(* IEC 61131-3 sources: BODAS-HelloWorld/st/bodas_rc18_12_40/plc_logic/application/02_easyconfig/dsm_easyconfig/structure (part 3) *)

(* ---- dfc_rbr_ina38scb-DFC_rbr_inA38SCB.st ---- *)
(* --- Interface --- *)
{attribute 'external_name' := 'cmp_rts_DFC_rbr_inA38SCB'}
TYPE DFC_rbr_inA38SCB : STRUCT
		DTC            : UDINT := 16#133100;
		DFCid          : UINT  := 257;
		debounceMethod : USINT := TIME_UP_DOWN;
	END_STRUCT
END_TYPE

(* ---- dfc_rbr_ina38scg-DFC_rbr_inA38SCG.st ---- *)
(* --- Interface --- *)
{attribute 'external_name' := 'cmp_rts_DFC_rbr_inA38SCG'}
TYPE DFC_rbr_inA38SCG : STRUCT
		DTC            : UDINT := 16#133200;
		DFCid          : UINT  := 258;
		debounceMethod : USINT := TIME_UP_DOWN;
	END_STRUCT
END_TYPE

(* ---- dfc_rbr_ina38shuntscb-DFC_rbr_inA38ShuntSCB.st ---- *)
(* --- Interface --- *)
{attribute 'external_name' := 'cmp_rts_DFC_rbr_inA38ShuntSCB'}
TYPE DFC_rbr_inA38ShuntSCB : STRUCT
		DTC            : UDINT := 16#133300;
		DFCid          : UINT  := 259;
		debounceMethod : USINT := TIME_UP_DOWN;
	END_STRUCT
END_TYPE

(* ---- dfc_rbr_ina39aicscb-DFC_rbr_inA39AicSCB.st ---- *)
(* --- Interface --- *)
{attribute 'external_name' := 'cmp_rts_DFC_rbr_inA39AicSCB'}
TYPE DFC_rbr_inA39AicSCB : STRUCT
		DTC            : UDINT := 16#133400;
		DFCid          : UINT  := 260;
		debounceMethod : USINT := TIME_UP_DOWN;
	END_STRUCT
END_TYPE

(* ---- dfc_rbr_ina39aicscg-DFC_rbr_inA39AicSCG.st ---- *)
(* --- Interface --- *)
{attribute 'external_name' := 'cmp_rts_DFC_rbr_inA39AicSCG'}
TYPE DFC_rbr_inA39AicSCG : STRUCT
		DTC            : UDINT := 16#133500;
		DFCid          : UINT  := 261;
		debounceMethod : USINT := TIME_UP_DOWN;
	END_STRUCT
END_TYPE

(* ---- dfc_rbr_ina39or-DFC_rbr_inA39OR.st ---- *)
(* --- Interface --- *)
{attribute 'external_name' := 'cmp_rts_DFC_rbr_inA39OR'}
TYPE DFC_rbr_inA39OR : STRUCT
		DTC            : UDINT := 16#133600;
		DFCid          : UINT  := 262;
		debounceMethod : USINT := TIME_UP_DOWN;
	END_STRUCT
END_TYPE

(* ---- dfc_rbr_ina39scb-DFC_rbr_inA39SCB.st ---- *)
(* --- Interface --- *)
{attribute 'external_name' := 'cmp_rts_DFC_rbr_inA39SCB'}
TYPE DFC_rbr_inA39SCB : STRUCT
		DTC            : UDINT := 16#133700;
		DFCid          : UINT  := 263;
		debounceMethod : USINT := TIME_UP_DOWN;
	END_STRUCT
END_TYPE

(* ---- dfc_rbr_ina39scg-DFC_rbr_inA39SCG.st ---- *)
(* --- Interface --- *)
{attribute 'external_name' := 'cmp_rts_DFC_rbr_inA39SCG'}
TYPE DFC_rbr_inA39SCG : STRUCT
		DTC            : UDINT := 16#133800;
		DFCid          : UINT  := 264;
		debounceMethod : USINT := TIME_UP_DOWN;
	END_STRUCT
END_TYPE

(* ---- dfc_rbr_ina39shuntscb-DFC_rbr_inA39ShuntSCB.st ---- *)
(* --- Interface --- *)
{attribute 'external_name' := 'cmp_rts_DFC_rbr_inA39ShuntSCB'}
TYPE DFC_rbr_inA39ShuntSCB : STRUCT
		DTC            : UDINT := 16#133900;
		DFCid          : UINT  := 265;
		debounceMethod : USINT := TIME_UP_DOWN;
	END_STRUCT
END_TYPE

(* ---- dfc_rbr_ina40or-DFC_rbr_inA40OR.st ---- *)
(* --- Interface --- *)
{attribute 'external_name' := 'cmp_rts_DFC_rbr_inA40OR'}
TYPE DFC_rbr_inA40OR : STRUCT
		DTC            : UDINT := 16#133A00;
		DFCid          : UINT  := 266;
		debounceMethod : USINT := TIME_UP_DOWN;
	END_STRUCT
END_TYPE

(* ---- dfc_rbr_ina40scb-DFC_rbr_inA40SCB.st ---- *)
(* --- Interface --- *)
{attribute 'external_name' := 'cmp_rts_DFC_rbr_inA40SCB'}
TYPE DFC_rbr_inA40SCB : STRUCT
		DTC            : UDINT := 16#133B00;
		DFCid          : UINT  := 267;
		debounceMethod : USINT := TIME_UP_DOWN;
	END_STRUCT
END_TYPE

(* ---- dfc_rbr_ina40scg-DFC_rbr_inA40SCG.st ---- *)
(* --- Interface --- *)
{attribute 'external_name' := 'cmp_rts_DFC_rbr_inA40SCG'}
TYPE DFC_rbr_inA40SCG : STRUCT
		DTC            : UDINT := 16#133C00;
		DFCid          : UINT  := 268;
		debounceMethod : USINT := TIME_UP_DOWN;
	END_STRUCT
END_TYPE

(* ---- dfc_rbr_ina41or-DFC_rbr_inA41OR.st ---- *)
(* --- Interface --- *)
{attribute 'external_name' := 'cmp_rts_DFC_rbr_inA41OR'}
TYPE DFC_rbr_inA41OR : STRUCT
		DTC            : UDINT := 16#133D00;
		DFCid          : UINT  := 269;
		debounceMethod : USINT := TIME_UP_DOWN;
	END_STRUCT
END_TYPE

(* ---- dfc_rbr_ina41scb-DFC_rbr_inA41SCB.st ---- *)
(* --- Interface --- *)
{attribute 'external_name' := 'cmp_rts_DFC_rbr_inA41SCB'}
TYPE DFC_rbr_inA41SCB : STRUCT
		DTC            : UDINT := 16#133E00;
		DFCid          : UINT  := 270;
		debounceMethod : USINT := TIME_UP_DOWN;
	END_STRUCT
END_TYPE

(* ---- dfc_rbr_ina41scg-DFC_rbr_inA41SCG.st ---- *)
(* --- Interface --- *)
{attribute 'external_name' := 'cmp_rts_DFC_rbr_inA41SCG'}
TYPE DFC_rbr_inA41SCG : STRUCT
		DTC            : UDINT := 16#133F00;
		DFCid          : UINT  := 271;
		debounceMethod : USINT := TIME_UP_DOWN;
	END_STRUCT
END_TYPE

(* ---- dfc_rbr_ina42or-DFC_rbr_inA42OR.st ---- *)
(* --- Interface --- *)
{attribute 'external_name' := 'cmp_rts_DFC_rbr_inA42OR'}
TYPE DFC_rbr_inA42OR : STRUCT
		DTC            : UDINT := 16#134000;
		DFCid          : UINT  := 272;
		debounceMethod : USINT := TIME_UP_DOWN;
	END_STRUCT
END_TYPE

(* ---- dfc_rbr_ina42scb-DFC_rbr_inA42SCB.st ---- *)
(* --- Interface --- *)
{attribute 'external_name' := 'cmp_rts_DFC_rbr_inA42SCB'}
TYPE DFC_rbr_inA42SCB : STRUCT
		DTC            : UDINT := 16#134100;
		DFCid          : UINT  := 273;
		debounceMethod : USINT := TIME_UP_DOWN;
	END_STRUCT
END_TYPE

(* ---- dfc_rbr_ina42scg-DFC_rbr_inA42SCG.st ---- *)
(* --- Interface --- *)
{attribute 'external_name' := 'cmp_rts_DFC_rbr_inA42SCG'}
TYPE DFC_rbr_inA42SCG : STRUCT
		DTC            : UDINT := 16#134200;
		DFCid          : UINT  := 274;
		debounceMethod : USINT := TIME_UP_DOWN;
	END_STRUCT
END_TYPE

(* ---- dfc_rbr_ina43aicscb-DFC_rbr_inA43AicSCB.st ---- *)
(* --- Interface --- *)
{attribute 'external_name' := 'cmp_rts_DFC_rbr_inA43AicSCB'}
TYPE DFC_rbr_inA43AicSCB : STRUCT
		DTC            : UDINT := 16#134300;
		DFCid          : UINT  := 275;
		debounceMethod : USINT := TIME_UP_DOWN;
	END_STRUCT
END_TYPE

(* ---- dfc_rbr_ina43aicscg-DFC_rbr_inA43AicSCG.st ---- *)
(* --- Interface --- *)
{attribute 'external_name' := 'cmp_rts_DFC_rbr_inA43AicSCG'}
TYPE DFC_rbr_inA43AicSCG : STRUCT
		DTC            : UDINT := 16#134400;
		DFCid          : UINT  := 276;
		debounceMethod : USINT := TIME_UP_DOWN;
	END_STRUCT
END_TYPE

(* ---- dfc_rbr_ina43or-DFC_rbr_inA43OR.st ---- *)
(* --- Interface --- *)
{attribute 'external_name' := 'cmp_rts_DFC_rbr_inA43OR'}
TYPE DFC_rbr_inA43OR : STRUCT
		DTC            : UDINT := 16#134500;
		DFCid          : UINT  := 277;
		debounceMethod : USINT := TIME_UP_DOWN;
	END_STRUCT
END_TYPE

(* ---- dfc_rbr_ina43scb-DFC_rbr_inA43SCB.st ---- *)
(* --- Interface --- *)
{attribute 'external_name' := 'cmp_rts_DFC_rbr_inA43SCB'}
TYPE DFC_rbr_inA43SCB : STRUCT
		DTC            : UDINT := 16#134600;
		DFCid          : UINT  := 278;
		debounceMethod : USINT := TIME_UP_DOWN;
	END_STRUCT
END_TYPE

(* ---- dfc_rbr_ina43scg-DFC_rbr_inA43SCG.st ---- *)
(* --- Interface --- *)
{attribute 'external_name' := 'cmp_rts_DFC_rbr_inA43SCG'}
TYPE DFC_rbr_inA43SCG : STRUCT
		DTC            : UDINT := 16#134700;
		DFCid          : UINT  := 279;
		debounceMethod : USINT := TIME_UP_DOWN;
	END_STRUCT
END_TYPE

(* ---- dfc_rbr_ina43shuntscb-DFC_rbr_inA43ShuntSCB.st ---- *)
(* --- Interface --- *)
{attribute 'external_name' := 'cmp_rts_DFC_rbr_inA43ShuntSCB'}
TYPE DFC_rbr_inA43ShuntSCB : STRUCT
		DTC            : UDINT := 16#134800;
		DFCid          : UINT  := 280;
		debounceMethod : USINT := TIME_UP_DOWN;
	END_STRUCT
END_TYPE

(* ---- dfc_rbr_ina44ol-DFC_rbr_inA44OL.st ---- *)
(* --- Interface --- *)
{attribute 'external_name' := 'cmp_rts_DFC_rbr_inA44OL'}
TYPE DFC_rbr_inA44OL : STRUCT
		DTC            : UDINT := 16#134900;
		DFCid          : UINT  := 281;
		debounceMethod : USINT := TIME_UP_DOWN;
	END_STRUCT
END_TYPE

(* ---- dfc_rbr_ina44scb-DFC_rbr_inA44SCB.st ---- *)
(* --- Interface --- *)
{attribute 'external_name' := 'cmp_rts_DFC_rbr_inA44SCB'}
TYPE DFC_rbr_inA44SCB : STRUCT
		DTC            : UDINT := 16#134A00;
		DFCid          : UINT  := 282;
		debounceMethod : USINT := TIME_UP_DOWN;
	END_STRUCT
END_TYPE

(* ---- dfc_rbr_ina44scg-DFC_rbr_inA44SCG.st ---- *)
(* --- Interface --- *)
{attribute 'external_name' := 'cmp_rts_DFC_rbr_inA44SCG'}
TYPE DFC_rbr_inA44SCG : STRUCT
		DTC            : UDINT := 16#134B00;
		DFCid          : UINT  := 283;
		debounceMethod : USINT := TIME_UP_DOWN;
	END_STRUCT
END_TYPE

(* ---- dfc_rbr_ina57or-DFC_rbr_inA57OR.st ---- *)
(* --- Interface --- *)
{attribute 'external_name' := 'cmp_rts_DFC_rbr_inA57OR'}
TYPE DFC_rbr_inA57OR : STRUCT
		DTC            : UDINT := 16#134C00;
		DFCid          : UINT  := 284;
		debounceMethod : USINT := TIME_UP_DOWN;
	END_STRUCT
END_TYPE

(* ---- dfc_rbr_ina57scb-DFC_rbr_inA57SCB.st ---- *)
(* --- Interface --- *)
{attribute 'external_name' := 'cmp_rts_DFC_rbr_inA57SCB'}
TYPE DFC_rbr_inA57SCB : STRUCT
		DTC            : UDINT := 16#134D00;
		DFCid          : UINT  := 285;
		debounceMethod : USINT := TIME_UP_DOWN;
	END_STRUCT
END_TYPE

(* ---- dfc_rbr_ina57scg-DFC_rbr_inA57SCG.st ---- *)
(* --- Interface --- *)
{attribute 'external_name' := 'cmp_rts_DFC_rbr_inA57SCG'}
TYPE DFC_rbr_inA57SCG : STRUCT
		DTC            : UDINT := 16#134E00;
		DFCid          : UINT  := 286;
		debounceMethod : USINT := TIME_UP_DOWN;
	END_STRUCT
END_TYPE

(* ---- dfc_rbr_ina59ol-DFC_rbr_inA59OL.st ---- *)
(* --- Interface --- *)
{attribute 'external_name' := 'cmp_rts_DFC_rbr_inA59OL'}
TYPE DFC_rbr_inA59OL : STRUCT
		DTC            : UDINT := 16#134F00;
		DFCid          : UINT  := 287;
		debounceMethod : USINT := TIME_UP_DOWN;
	END_STRUCT
END_TYPE

(* ---- dfc_rbr_ina59scb-DFC_rbr_inA59SCB.st ---- *)
(* --- Interface --- *)
{attribute 'external_name' := 'cmp_rts_DFC_rbr_inA59SCB'}
TYPE DFC_rbr_inA59SCB : STRUCT
		DTC            : UDINT := 16#135000;
		DFCid          : UINT  := 288;
		debounceMethod : USINT := TIME_UP_DOWN;
	END_STRUCT
END_TYPE

(* ---- dfc_rbr_ina59scg-DFC_rbr_inA59SCG.st ---- *)
(* --- Interface --- *)
{attribute 'external_name' := 'cmp_rts_DFC_rbr_inA59SCG'}
TYPE DFC_rbr_inA59SCG : STRUCT
		DTC            : UDINT := 16#135100;
		DFCid          : UINT  := 289;
		debounceMethod : USINT := TIME_UP_DOWN;
	END_STRUCT
END_TYPE

(* ---- dfc_rbr_inai-DFC_rbr_inAi.st ---- *)
(* --- Interface --- *)
{attribute 'external_name' := 'cmp_rts_DFC_rbr_inAi'}
TYPE DFC_rbr_inAi : STRUCT
		DTC            : UDINT := 16#038000;
		DFCid          : UINT  := 882;
		debounceMethod : USINT := NO_DEBOUNCE;
	END_STRUCT
END_TYPE

(* ---- dfc_rbr_inaic-DFC_rbr_inAic.st ---- *)
(* --- Interface --- *)
{attribute 'external_name' := 'cmp_rts_DFC_rbr_inAic'}
TYPE DFC_rbr_inAic : STRUCT
		DTC            : UDINT := 16#038100;
		DFCid          : UINT  := 883;
		debounceMethod : USINT := NO_DEBOUNCE;
	END_STRUCT
END_TYPE

(* ---- dfc_rbr_inaiccfg-DFC_rbr_inAicCfg.st ---- *)
(* --- Interface --- *)
{attribute 'external_name' := 'cmp_rts_DFC_rbr_inAicCfg'}
TYPE DFC_rbr_inAicCfg : STRUCT
		DTC            : UDINT := 16#038200;
		DFCid          : UINT  := 884;
		debounceMethod : USINT := NO_DEBOUNCE;
	END_STRUCT
END_TYPE

(* ---- dfc_rbr_inaicgetstatus-DFC_rbr_inAicGetStatus.st ---- *)
(* --- Interface --- *)
{attribute 'external_name' := 'cmp_rts_DFC_rbr_inAicGetStatus'}
TYPE DFC_rbr_inAicGetStatus : STRUCT
		DTC            : UDINT := 16#038D00;
		DFCid          : UINT  := 885;
		debounceMethod : USINT := NO_DEBOUNCE;
	END_STRUCT
END_TYPE

(* ---- dfc_rbr_inaid-DFC_rbr_inAid.st ---- *)
(* --- Interface --- *)
{attribute 'external_name' := 'cmp_rts_DFC_rbr_inAid'}
TYPE DFC_rbr_inAid : STRUCT
		DTC            : UDINT := 16#038300;
		DFCid          : UINT  := 886;
		debounceMethod : USINT := NO_DEBOUNCE;
	END_STRUCT
END_TYPE

(* ---- dfc_rbr_inaidcfg-DFC_rbr_inAidCfg.st ---- *)
(* --- Interface --- *)
{attribute 'external_name' := 'cmp_rts_DFC_rbr_inAidCfg'}
TYPE DFC_rbr_inAidCfg : STRUCT
		DTC            : UDINT := 16#038400;
		DFCid          : UINT  := 887;
		debounceMethod : USINT := NO_DEBOUNCE;
	END_STRUCT
END_TYPE

(* ---- dfc_rbr_inaiv-DFC_rbr_inAiv.st ---- *)
(* --- Interface --- *)
{attribute 'external_name' := 'cmp_rts_DFC_rbr_inAiv'}
TYPE DFC_rbr_inAiv : STRUCT
		DTC            : UDINT := 16#038500;
		DFCid          : UINT  := 888;
		debounceMethod : USINT := NO_DEBOUNCE;
	END_STRUCT
END_TYPE

(* ---- dfc_rbr_inaivcfg-DFC_rbr_inAivCfg.st ---- *)
(* --- Interface --- *)
{attribute 'external_name' := 'cmp_rts_DFC_rbr_inAivCfg'}
TYPE DFC_rbr_inAivCfg : STRUCT
		DTC            : UDINT := 16#038600;
		DFCid          : UINT  := 889;
		debounceMethod : USINT := NO_DEBOUNCE;
	END_STRUCT
END_TYPE

(* ---- dfc_rbr_inaivgetstatus-DFC_rbr_inAivGetStatus.st ---- *)
(* --- Interface --- *)
{attribute 'external_name' := 'cmp_rts_DFC_rbr_inAivGetStatus'}
TYPE DFC_rbr_inAivGetStatus : STRUCT
		DTC            : UDINT := 16#038C00;
		DFCid          : UINT  := 890;
		debounceMethod : USINT := NO_DEBOUNCE;
	END_STRUCT
END_TYPE

(* ---- dfc_rbr_indi-DFC_rbr_inDi.st ---- *)
(* --- Interface --- *)
{attribute 'external_name' := 'cmp_rts_DFC_rbr_inDi'}
TYPE DFC_rbr_inDi : STRUCT
		DTC            : UDINT := 16#038700;
		DFCid          : UINT  := 891;
		debounceMethod : USINT := NO_DEBOUNCE;
	END_STRUCT
END_TYPE

(* ---- dfc_rbr_infi-DFC_rbr_inFi.st ---- *)
(* --- Interface --- *)
{attribute 'external_name' := 'cmp_rts_DFC_rbr_inFi'}
TYPE DFC_rbr_inFi : STRUCT
		DTC            : UDINT := 16#038800;
		DFCid          : UINT  := 892;
		debounceMethod : USINT := NO_DEBOUNCE;
	END_STRUCT
END_TYPE

(* ---- dfc_rbr_infi_buffered-DFC_rbr_inFi_Buffered.st ---- *)
(* --- Interface --- *)
{attribute 'external_name' := 'cmp_rts_DFC_rbr_inFi_Buffered'}
TYPE DFC_rbr_inFi_Buffered : STRUCT
		DTC            : UDINT := 16#135200;
		DFCid          : UINT  := 895;
		debounceMethod : USINT := NO_DEBOUNCE;
	END_STRUCT
END_TYPE

(* ---- dfc_rbr_inficfg-DFC_rbr_inFiCfg.st ---- *)
(* --- Interface --- *)
{attribute 'external_name' := 'cmp_rts_DFC_rbr_inFiCfg'}
TYPE DFC_rbr_inFiCfg : STRUCT
		DTC            : UDINT := 16#038900;
		DFCid          : UINT  := 893;
		debounceMethod : USINT := NO_DEBOUNCE;
	END_STRUCT
END_TYPE

(* ---- dfc_rbr_infigetstatus-DFC_rbr_inFiGetStatus.st ---- *)
(* --- Interface --- *)
{attribute 'external_name' := 'cmp_rts_DFC_rbr_inFiGetStatus'}
TYPE DFC_rbr_inFiGetStatus : STRUCT
		DTC            : UDINT := 16#038F00;
		DFCid          : UINT  := 894;
		debounceMethod : USINT := NO_DEBOUNCE;
	END_STRUCT
END_TYPE

(* ---- dfc_rbr_ink10or-DFC_rbr_inK10OR.st ---- *)
(* --- Interface --- *)
{attribute 'external_name' := 'cmp_rts_DFC_rbr_inK10OR'}
TYPE DFC_rbr_inK10OR : STRUCT
		DTC            : UDINT := 16#030100;
		DFCid          : UINT  := 290;
		debounceMethod : USINT := TIME_UP_DOWN;
	END_STRUCT
END_TYPE

(* ---- dfc_rbr_ink10scb-DFC_rbr_inK10SCB.st ---- *)
(* --- Interface --- *)
{attribute 'external_name' := 'cmp_rts_DFC_rbr_inK10SCB'}
TYPE DFC_rbr_inK10SCB : STRUCT
		DTC            : UDINT := 16#030200;
		DFCid          : UINT  := 291;
		debounceMethod : USINT := TIME_UP_DOWN;
	END_STRUCT
END_TYPE

(* ---- dfc_rbr_ink10scg-DFC_rbr_inK10SCG.st ---- *)
(* --- Interface --- *)
{attribute 'external_name' := 'cmp_rts_DFC_rbr_inK10SCG'}
TYPE DFC_rbr_inK10SCG : STRUCT
		DTC            : UDINT := 16#030300;
		DFCid          : UINT  := 292;
		debounceMethod : USINT := TIME_UP_DOWN;
	END_STRUCT
END_TYPE

(* ---- dfc_rbr_ink11or-DFC_rbr_inK11OR.st ---- *)
(* --- Interface --- *)
{attribute 'external_name' := 'cmp_rts_DFC_rbr_inK11OR'}
TYPE DFC_rbr_inK11OR : STRUCT
		DTC            : UDINT := 16#03A200;
		DFCid          : UINT  := 293;
		debounceMethod : USINT := TIME_UP_DOWN;
	END_STRUCT
END_TYPE

(* ---- dfc_rbr_ink11scb-DFC_rbr_inK11SCB.st ---- *)
(* --- Interface --- *)
{attribute 'external_name' := 'cmp_rts_DFC_rbr_inK11SCB'}
TYPE DFC_rbr_inK11SCB : STRUCT
		DTC            : UDINT := 16#03A300;
		DFCid          : UINT  := 294;
		debounceMethod : USINT := TIME_UP_DOWN;
	END_STRUCT
END_TYPE

(* ---- dfc_rbr_ink11scg-DFC_rbr_inK11SCG.st ---- *)
(* --- Interface --- *)
{attribute 'external_name' := 'cmp_rts_DFC_rbr_inK11SCG'}
TYPE DFC_rbr_inK11SCG : STRUCT
		DTC            : UDINT := 16#03A400;
		DFCid          : UINT  := 295;
		debounceMethod : USINT := TIME_UP_DOWN;
	END_STRUCT
END_TYPE

(* ---- dfc_rbr_ink30aicscb-DFC_rbr_inK30AicSCB.st ---- *)
(* --- Interface --- *)
{attribute 'external_name' := 'cmp_rts_DFC_rbr_inK30AicSCB'}
TYPE DFC_rbr_inK30AicSCB : STRUCT
		DTC            : UDINT := 16#03A500;
		DFCid          : UINT  := 296;
		debounceMethod : USINT := TIME_UP_DOWN;
	END_STRUCT
END_TYPE

(* ---- dfc_rbr_ink30aicscg-DFC_rbr_inK30AicSCG.st ---- *)
(* --- Interface --- *)
{attribute 'external_name' := 'cmp_rts_DFC_rbr_inK30AicSCG'}
TYPE DFC_rbr_inK30AicSCG : STRUCT
		DTC            : UDINT := 16#03A600;
		DFCid          : UINT  := 297;
		debounceMethod : USINT := TIME_UP_DOWN;
	END_STRUCT
END_TYPE

(* ---- dfc_rbr_ink30or-DFC_rbr_inK30OR.st ---- *)
(* --- Interface --- *)
{attribute 'external_name' := 'cmp_rts_DFC_rbr_inK30OR'}
TYPE DFC_rbr_inK30OR : STRUCT
		DTC            : UDINT := 16#03A700;
		DFCid          : UINT  := 298;
		debounceMethod : USINT := TIME_UP_DOWN;
	END_STRUCT
END_TYPE

(* ---- dfc_rbr_ink30scb-DFC_rbr_inK30SCB.st ---- *)
(* --- Interface --- *)
{attribute 'external_name' := 'cmp_rts_DFC_rbr_inK30SCB'}
TYPE DFC_rbr_inK30SCB : STRUCT
		DTC            : UDINT := 16#03A800;
		DFCid          : UINT  := 299;
		debounceMethod : USINT := TIME_UP_DOWN;
	END_STRUCT
END_TYPE

(* ---- dfc_rbr_ink30scg-DFC_rbr_inK30SCG.st ---- *)
(* --- Interface --- *)
{attribute 'external_name' := 'cmp_rts_DFC_rbr_inK30SCG'}
TYPE DFC_rbr_inK30SCG : STRUCT
		DTC            : UDINT := 16#03A900;
		DFCid          : UINT  := 300;
		debounceMethod : USINT := TIME_UP_DOWN;
	END_STRUCT
END_TYPE

(* ---- dfc_rbr_ink30shuntscb-DFC_rbr_inK30ShuntSCB.st ---- *)
(* --- Interface --- *)
{attribute 'external_name' := 'cmp_rts_DFC_rbr_inK30ShuntSCB'}
TYPE DFC_rbr_inK30ShuntSCB : STRUCT
		DTC            : UDINT := 16#03AA00;
		DFCid          : UINT  := 301;
		debounceMethod : USINT := TIME_UP_DOWN;
	END_STRUCT
END_TYPE

(* ---- dfc_rbr_ink31or-DFC_rbr_inK31OR.st ---- *)
(* --- Interface --- *)
{attribute 'external_name' := 'cmp_rts_DFC_rbr_inK31OR'}
TYPE DFC_rbr_inK31OR : STRUCT
		DTC            : UDINT := 16#03AB00;
		DFCid          : UINT  := 302;
		debounceMethod : USINT := TIME_UP_DOWN;
	END_STRUCT
END_TYPE

(* ---- dfc_rbr_ink31scb-DFC_rbr_inK31SCB.st ---- *)
(* --- Interface --- *)
{attribute 'external_name' := 'cmp_rts_DFC_rbr_inK31SCB'}
TYPE DFC_rbr_inK31SCB : STRUCT
		DTC            : UDINT := 16#03AC00;
		DFCid          : UINT  := 303;
		debounceMethod : USINT := TIME_UP_DOWN;
	END_STRUCT
END_TYPE

(* ---- dfc_rbr_ink31scg-DFC_rbr_inK31SCG.st ---- *)
(* --- Interface --- *)
{attribute 'external_name' := 'cmp_rts_DFC_rbr_inK31SCG'}
TYPE DFC_rbr_inK31SCG : STRUCT
		DTC            : UDINT := 16#03AD00;
		DFCid          : UINT  := 304;
		debounceMethod : USINT := TIME_UP_DOWN;
	END_STRUCT
END_TYPE

(* ---- dfc_rbr_ink32or-DFC_rbr_inK32OR.st ---- *)
(* --- Interface --- *)
{attribute 'external_name' := 'cmp_rts_DFC_rbr_inK32OR'}
TYPE DFC_rbr_inK32OR : STRUCT
		DTC            : UDINT := 16#03AE00;
		DFCid          : UINT  := 305;
		debounceMethod : USINT := TIME_UP_DOWN;
	END_STRUCT
END_TYPE

(* ---- dfc_rbr_ink32scb-DFC_rbr_inK32SCB.st ---- *)
(* --- Interface --- *)
{attribute 'external_name' := 'cmp_rts_DFC_rbr_inK32SCB'}
TYPE DFC_rbr_inK32SCB : STRUCT
		DTC            : UDINT := 16#03AF00;
		DFCid          : UINT  := 306;
		debounceMethod : USINT := TIME_UP_DOWN;
	END_STRUCT
END_TYPE

(* ---- dfc_rbr_ink32scg-DFC_rbr_inK32SCG.st ---- *)
(* --- Interface --- *)
{attribute 'external_name' := 'cmp_rts_DFC_rbr_inK32SCG'}
TYPE DFC_rbr_inK32SCG : STRUCT
		DTC            : UDINT := 16#03B000;
		DFCid          : UINT  := 307;
		debounceMethod : USINT := TIME_UP_DOWN;
	END_STRUCT
END_TYPE

(* ---- dfc_rbr_ink33or-DFC_rbr_inK33OR.st ---- *)
(* --- Interface --- *)
{attribute 'external_name' := 'cmp_rts_DFC_rbr_inK33OR'}
TYPE DFC_rbr_inK33OR : STRUCT
		DTC            : UDINT := 16#03B100;
		DFCid          : UINT  := 308;
		debounceMethod : USINT := TIME_UP_DOWN;
	END_STRUCT
END_TYPE

(* ---- dfc_rbr_ink33scb-DFC_rbr_inK33SCB.st ---- *)
(* --- Interface --- *)
{attribute 'external_name' := 'cmp_rts_DFC_rbr_inK33SCB'}
TYPE DFC_rbr_inK33SCB : STRUCT
		DTC            : UDINT := 16#03B200;
		DFCid          : UINT  := 309;
		debounceMethod : USINT := TIME_UP_DOWN;
	END_STRUCT
END_TYPE

(* ---- dfc_rbr_ink33scg-DFC_rbr_inK33SCG.st ---- *)
(* --- Interface --- *)
{attribute 'external_name' := 'cmp_rts_DFC_rbr_inK33SCG'}
TYPE DFC_rbr_inK33SCG : STRUCT
		DTC            : UDINT := 16#03B300;
		DFCid          : UINT  := 310;
		debounceMethod : USINT := TIME_UP_DOWN;
	END_STRUCT
END_TYPE

(* ---- dfc_rbr_ink34or-DFC_rbr_inK34OR.st ---- *)
(* --- Interface --- *)
{attribute 'external_name' := 'cmp_rts_DFC_rbr_inK34OR'}
TYPE DFC_rbr_inK34OR : STRUCT
		DTC            : UDINT := 16#03B400;
		DFCid          : UINT  := 311;
		debounceMethod : USINT := TIME_UP_DOWN;
	END_STRUCT
END_TYPE

(* ---- dfc_rbr_ink34scb-DFC_rbr_inK34SCB.st ---- *)
(* --- Interface --- *)
{attribute 'external_name' := 'cmp_rts_DFC_rbr_inK34SCB'}
TYPE DFC_rbr_inK34SCB : STRUCT
		DTC            : UDINT := 16#03B500;
		DFCid          : UINT  := 312;
		debounceMethod : USINT := TIME_UP_DOWN;
	END_STRUCT
END_TYPE

(* ---- dfc_rbr_ink34scg-DFC_rbr_inK34SCG.st ---- *)
(* --- Interface --- *)
{attribute 'external_name' := 'cmp_rts_DFC_rbr_inK34SCG'}
TYPE DFC_rbr_inK34SCG : STRUCT
		DTC            : UDINT := 16#03B600;
		DFCid          : UINT  := 313;
		debounceMethod : USINT := TIME_UP_DOWN;
	END_STRUCT
END_TYPE

(* ---- dfc_rbr_ink35or-DFC_rbr_inK35OR.st ---- *)
(* --- Interface --- *)
{attribute 'external_name' := 'cmp_rts_DFC_rbr_inK35OR'}
TYPE DFC_rbr_inK35OR : STRUCT
		DTC            : UDINT := 16#03B700;
		DFCid          : UINT  := 314;
		debounceMethod : USINT := TIME_UP_DOWN;
	END_STRUCT
END_TYPE

(* ---- dfc_rbr_ink35scb-DFC_rbr_inK35SCB.st ---- *)
(* --- Interface --- *)
{attribute 'external_name' := 'cmp_rts_DFC_rbr_inK35SCB'}
TYPE DFC_rbr_inK35SCB : STRUCT
		DTC            : UDINT := 16#03B800;
		DFCid          : UINT  := 315;
		debounceMethod : USINT := TIME_UP_DOWN;
	END_STRUCT
END_TYPE

(* ---- dfc_rbr_ink35scg-DFC_rbr_inK35SCG.st ---- *)
(* --- Interface --- *)
{attribute 'external_name' := 'cmp_rts_DFC_rbr_inK35SCG'}
TYPE DFC_rbr_inK35SCG : STRUCT
		DTC            : UDINT := 16#03B900;
		DFCid          : UINT  := 316;
		debounceMethod : USINT := TIME_UP_DOWN;
	END_STRUCT
END_TYPE

(* ---- dfc_rbr_ink36or-DFC_rbr_inK36OR.st ---- *)
(* --- Interface --- *)
{attribute 'external_name' := 'cmp_rts_DFC_rbr_inK36OR'}
TYPE DFC_rbr_inK36OR : STRUCT
		DTC            : UDINT := 16#030400;
		DFCid          : UINT  := 317;
		debounceMethod : USINT := TIME_UP_DOWN;
	END_STRUCT
END_TYPE

(* ---- dfc_rbr_ink36scb-DFC_rbr_inK36SCB.st ---- *)
(* --- Interface --- *)
{attribute 'external_name' := 'cmp_rts_DFC_rbr_inK36SCB'}
TYPE DFC_rbr_inK36SCB : STRUCT
		DTC            : UDINT := 16#030500;
		DFCid          : UINT  := 318;
		debounceMethod : USINT := TIME_UP_DOWN;
	END_STRUCT
END_TYPE

(* ---- dfc_rbr_ink36scg-DFC_rbr_inK36SCG.st ---- *)
(* --- Interface --- *)
{attribute 'external_name' := 'cmp_rts_DFC_rbr_inK36SCG'}
TYPE DFC_rbr_inK36SCG : STRUCT
		DTC            : UDINT := 16#030600;
		DFCid          : UINT  := 319;
		debounceMethod : USINT := TIME_UP_DOWN;
	END_STRUCT
END_TYPE

(* ---- dfc_rbr_ink37aicscb-DFC_rbr_inK37AicSCB.st ---- *)
(* --- Interface --- *)
{attribute 'external_name' := 'cmp_rts_DFC_rbr_inK37AicSCB'}
TYPE DFC_rbr_inK37AicSCB : STRUCT
		DTC            : UDINT := 16#030700;
		DFCid          : UINT  := 320;
		debounceMethod : USINT := TIME_UP_DOWN;
	END_STRUCT
END_TYPE

(* ---- dfc_rbr_ink37aicscg-DFC_rbr_inK37AicSCG.st ---- *)
(* --- Interface --- *)
{attribute 'external_name' := 'cmp_rts_DFC_rbr_inK37AicSCG'}
TYPE DFC_rbr_inK37AicSCG : STRUCT
		DTC            : UDINT := 16#030800;
		DFCid          : UINT  := 321;
		debounceMethod : USINT := TIME_UP_DOWN;
	END_STRUCT
END_TYPE

(* ---- dfc_rbr_ink37or-DFC_rbr_inK37OR.st ---- *)
(* --- Interface --- *)
{attribute 'external_name' := 'cmp_rts_DFC_rbr_inK37OR'}
TYPE DFC_rbr_inK37OR : STRUCT
		DTC            : UDINT := 16#030900;
		DFCid          : UINT  := 322;
		debounceMethod : USINT := TIME_UP_DOWN;
	END_STRUCT
END_TYPE

(* ---- dfc_rbr_ink37scb-DFC_rbr_inK37SCB.st ---- *)
(* --- Interface --- *)
{attribute 'external_name' := 'cmp_rts_DFC_rbr_inK37SCB'}
TYPE DFC_rbr_inK37SCB : STRUCT
		DTC            : UDINT := 16#030A00;
		DFCid          : UINT  := 323;
		debounceMethod : USINT := TIME_UP_DOWN;
	END_STRUCT
END_TYPE

(* ---- dfc_rbr_ink37scg-DFC_rbr_inK37SCG.st ---- *)
(* --- Interface --- *)
{attribute 'external_name' := 'cmp_rts_DFC_rbr_inK37SCG'}
TYPE DFC_rbr_inK37SCG : STRUCT
		DTC            : UDINT := 16#030B00;
		DFCid          : UINT  := 324;
		debounceMethod : USINT := TIME_UP_DOWN;
	END_STRUCT
END_TYPE

(* ---- dfc_rbr_ink37shuntscb-DFC_rbr_inK37ShuntSCB.st ---- *)
(* --- Interface --- *)
{attribute 'external_name' := 'cmp_rts_DFC_rbr_inK37ShuntSCB'}
TYPE DFC_rbr_inK37ShuntSCB : STRUCT
		DTC            : UDINT := 16#030C00;
		DFCid          : UINT  := 325;
		debounceMethod : USINT := TIME_UP_DOWN;
	END_STRUCT
END_TYPE

(* ---- dfc_rbr_ink38aicscb-DFC_rbr_inK38AicSCB.st ---- *)
(* --- Interface --- *)
{attribute 'external_name' := 'cmp_rts_DFC_rbr_inK38AicSCB'}
TYPE DFC_rbr_inK38AicSCB : STRUCT
		DTC            : UDINT := 16#03BA00;
		DFCid          : UINT  := 326;
		debounceMethod : USINT := TIME_UP_DOWN;
	END_STRUCT
END_TYPE

(* ---- dfc_rbr_ink38aicscg-DFC_rbr_inK38AicSCG.st ---- *)
(* --- Interface --- *)
{attribute 'external_name' := 'cmp_rts_DFC_rbr_inK38AicSCG'}
TYPE DFC_rbr_inK38AicSCG : STRUCT
		DTC            : UDINT := 16#03BB00;
		DFCid          : UINT  := 327;
		debounceMethod : USINT := TIME_UP_DOWN;
	END_STRUCT
END_TYPE

(* ---- dfc_rbr_ink38or-DFC_rbr_inK38OR.st ---- *)
(* --- Interface --- *)
{attribute 'external_name' := 'cmp_rts_DFC_rbr_inK38OR'}
TYPE DFC_rbr_inK38OR : STRUCT
		DTC            : UDINT := 16#030D00;
		DFCid          : UINT  := 328;
		debounceMethod : USINT := TIME_UP_DOWN;
	END_STRUCT
END_TYPE

(* ---- dfc_rbr_ink38scb-DFC_rbr_inK38SCB.st ---- *)
(* --- Interface --- *)
{attribute 'external_name' := 'cmp_rts_DFC_rbr_inK38SCB'}
TYPE DFC_rbr_inK38SCB : STRUCT
		DTC            : UDINT := 16#030E00;
		DFCid          : UINT  := 329;
		debounceMethod : USINT := TIME_UP_DOWN;
	END_STRUCT
END_TYPE

(* ---- dfc_rbr_ink38scg-DFC_rbr_inK38SCG.st ---- *)
(* --- Interface --- *)
{attribute 'external_name' := 'cmp_rts_DFC_rbr_inK38SCG'}
TYPE DFC_rbr_inK38SCG : STRUCT
		DTC            : UDINT := 16#030F00;
		DFCid          : UINT  := 330;
		debounceMethod : USINT := TIME_UP_DOWN;
	END_STRUCT
END_TYPE

(* ---- dfc_rbr_ink38shuntscb-DFC_rbr_inK38ShuntSCB.st ---- *)
(* --- Interface --- *)
{attribute 'external_name' := 'cmp_rts_DFC_rbr_inK38ShuntSCB'}
TYPE DFC_rbr_inK38ShuntSCB : STRUCT
		DTC            : UDINT := 16#03BC00;
		DFCid          : UINT  := 331;
		debounceMethod : USINT := TIME_UP_DOWN;
	END_STRUCT
END_TYPE

(* ---- dfc_rbr_ink39aicscb-DFC_rbr_inK39AicSCB.st ---- *)
(* --- Interface --- *)
{attribute 'external_name' := 'cmp_rts_DFC_rbr_inK39AicSCB'}
TYPE DFC_rbr_inK39AicSCB : STRUCT
		DTC            : UDINT := 16#03BD00;
		DFCid          : UINT  := 332;
		debounceMethod : USINT := TIME_UP_DOWN;
	END_STRUCT
END_TYPE

(* ---- dfc_rbr_ink39aicscg-DFC_rbr_inK39AicSCG.st ---- *)
(* --- Interface --- *)
{attribute 'external_name' := 'cmp_rts_DFC_rbr_inK39AicSCG'}
TYPE DFC_rbr_inK39AicSCG : STRUCT
		DTC            : UDINT := 16#03BE00;
		DFCid          : UINT  := 333;
		debounceMethod : USINT := TIME_UP_DOWN;
	END_STRUCT
END_TYPE
